// Implicitly generated code : DO NOT EDIT
FUNCTION CheckBounds : DINT
VAR_INPUT
	index, lower, upper: DINT;
END_VAR
VAR_STAT
	nIndexOverflow : UDINT;
	nIndexUnderflow : UDINT;
END_VAR

// Implicitly generated code: Only an implementation suggestion
{noflow}
IF  index < lower THEN
	nIndexUnderflow := nIndexUnderflow + 1;
	CheckBounds := lower;
ELSIF  index > upper THEN
	nIndexOverflow := nIndexOverflow + 1;
	CheckBounds := upper;
ELSE  
	CheckBounds := index;
END_IF

END_FUNCTION

(* stored: Version 1.1.0.1, ProductVersion 3.1.4026.18
   POU CheckBounds: Id {990c4c5c-1e70-4092-9aed-cf5aa9d669b5}, SpecialFunc CheckBounds *)
